# EPICS autosave request: iocs/ad/mythen-ioc/db/mythen_settings.req
file "ADBase_settings.req", P=$(P), R=$(R)
# C also includes NDFile_settings.req and names NumCycles; mythen.template
# has neither record, so each save reported 27 PVs unconnected.
$(P)$(R)Setting
$(P)$(R)BeamEnergy
$(P)$(R)ThresholdEnergy
$(P)$(R)UseFlatField
$(P)$(R)UseCountRate
$(P)$(R)Tau
$(P)$(R)UseBadChanIntrpl
$(P)$(R)BitDepth
$(P)$(R)TriggerMode
$(P)$(R)DelayTime
$(P)$(R)UseGates
$(P)$(R)NumGates
$(P)$(R)NumFrames
$(P)$(R)ReadMode
